// TIA Portal V21 export
DATA_BLOCK "IDB_LadBoxes"   // DB20
// stored: InstanceOfName FB_LadBoxes, InstanceOfType FB
"FB_LadBoxes"
   // VAR_INPUT
   //    Start : Bool;
   //    InValue : Int;
   //    Limit : Int;
   // END_VAR
   // VAR_OUTPUT
   //    Delayed : Bool;
   //    Copy : Int;
   //    Sum : Int;
   //    IsEqual : Bool;
   //    IsGreater : Bool;
   //    IsLessEqual : Bool;
   //    Average : Real;
   //    SectionsOk : Bool;
   //    Skipped : Bool;
   //    AfterJump : Bool;
   // END_VAR
   // VAR
   //    Delay { S7_SetPoint := 'True'} : TON_TIME;
   //    DelayElapsed : Time;
   //    Sections { S7_SetPoint := 'True'} : "FB_SclSections";
   //    Values : Array[0..9] of Real;
   //    SectionsBusy : Bool;
   //    SectionsSteps : Int;
   //    Setpoint : Real;
   // END_VAR
BEGIN
END_DATA_BLOCK
